// TIA Portal V20 export
Screen "Sew_APC"  1276x673
  ScreenItem "Rectangle_3" at 194,365 size 865x300  Type=HmiRectangle
  ScreenItem "Rectangle_1" at 195,113 size 866x250  Type=HmiRectangle
  ScreenItem "Title_ScreenOverview_X390_Y2" at 390,7 size 510x57  Type=HmiTextBox
  ScreenItem "符号 IO 域_7" at 479,72 size 290x38  Type=HmiSymbolicIOField
  ScreenItem "Text field_1" at 194,113 size 866x31  Type=HmiTextBox
  ScreenItem "按钮_2" at 279,171 size 140x60  Type=HmiButton
  ScreenItem "permanentareaborderrectangle" at 0,0 size 0x0  Type=HmiRectangle
  ScreenItem "Line_Header_X0_Y64" at 0,65 size 1276x0  Type=HmiLine
  ScreenItem "Button_Back" at 2,2 size 90x60  Type=HmiButton
  ScreenItem "Frame_SendToDrive_1" at 201,369 size 199x294  Type=HmiRectangle
  ScreenItem "Text_ConrolDataToDrive_1" at 205,373 size 148x21  Type=HmiTextBox
  ScreenItem "Text_DigitalOutputs_33" at 229,397 size 146x16  Type=HmiTextBox
  ScreenItem "Text_DigitalOutputs_34" at 229,412 size 124x16  Type=HmiTextBox
  ScreenItem "Text_DigitalOutputs_35" at 229,428 size 124x16  Type=HmiTextBox
  ScreenItem "Text_DigitalOutputs_40" at 229,444 size 124x16  Type=HmiTextBox
  ScreenItem "Text_DigitalOutputs_36" at 229,460 size 124x16  Type=HmiTextBox
  ScreenItem "Text_DigitalOutputs_37" at 229,476 size 124x16  Type=HmiTextBox
  ScreenItem "Text_DigitalOutputs_24" at 229,492 size 124x16  Type=HmiTextBox
  ScreenItem "Text_DigitalOutputs_38" at 229,508 size 124x16  Type=HmiTextBox
  ScreenItem "Text_DigitalOutputs_25" at 229,524 size 124x16  Type=HmiTextBox
  ScreenItem "Text_DigitalOutputs_39" at 229,540 size 124x16  Type=HmiTextBox
  ScreenItem "Text_DigitalOutputs_26" at 229,556 size 124x16  Type=HmiTextBox
  ScreenItem "Text_DigitalOutputs_1" at 229,572 size 124x16  Type=HmiTextBox
  ScreenItem "Text_DigitalOutputs_28" at 229,588 size 161x16  Type=HmiTextBox
  ScreenItem "Text_DigitalOutputs_30" at 229,604 size 124x16  Type=HmiTextBox
  ScreenItem "Text_DigitalOutputs_31" at 229,620 size 124x16  Type=HmiTextBox
  ScreenItem "Text_DigitalOutputs_32" at 229,636 size 124x16  Type=HmiTextBox
  ScreenItem "LED_1_Left_23" at 0,0 size 100x30  Type=HmiCircle
  ScreenItem "LED_1_Left_22" at 0,0 size 100x30  Type=HmiCircle
  ScreenItem "LED_1_Left_21" at 0,0 size 100x30  Type=HmiCircle
  ScreenItem "LED_1_Left_20" at 0,0 size 100x30  Type=HmiCircle
  ScreenItem "LED_1_Left_19" at 0,0 size 100x30  Type=HmiCircle
  ScreenItem "LED_1_Left_18" at 0,0 size 100x30  Type=HmiCircle
  ScreenItem "LED_1_Left_40" at 0,0 size 100x30  Type=HmiCircle
  ScreenItem "LED_1_Left_17" at 0,0 size 100x30  Type=HmiCircle
  ScreenItem "LED_1_Left_39" at 0,0 size 100x30  Type=HmiCircle
  ScreenItem "LED_1_Left_16" at 0,0 size 100x30  Type=HmiCircle
  ScreenItem "LED_1_Left_38" at 0,0 size 100x30  Type=HmiCircle
  ScreenItem "LED_1_Left_37" at 0,0 size 100x30  Type=HmiCircle
  ScreenItem "LED_1_Left_36" at 0,0 size 100x30  Type=HmiCircle
  ScreenItem "LED_1_Left_35" at 0,0 size 100x30  Type=HmiCircle
  ScreenItem "LED_1_Left_34" at 0,0 size 100x30  Type=HmiCircle
  ScreenItem "LED_1_Left_33" at 0,0 size 100x30  Type=HmiCircle
  ScreenItem "Frame_SendToDrive_3" at 405,369 size 199x294  Type=HmiRectangle
  ScreenItem "Text_ConrolDataToDrive_2" at 407,372 size 148x23  Type=HmiTextBox
  ScreenItem "Text_DigitalOutputs_2" at 426,395 size 124x20  Type=HmiTextBox
  ScreenItem "Text_DigitalOutputs_3" at 426,410 size 124x20  Type=HmiTextBox
  ScreenItem "Text_DigitalOutputs_4" at 426,426 size 124x20  Type=HmiTextBox
  ScreenItem "Text_DigitalOutputs_5" at 426,458 size 124x20  Type=HmiTextBox
  ScreenItem "Text_DigitalOutputs_6" at 426,474 size 124x20  Type=HmiTextBox
  ScreenItem "Text_DigitalOutputs_7" at 426,490 size 158x20  Type=HmiTextBox
  ScreenItem "Text_DigitalOutputs_8" at 426,506 size 124x20  Type=HmiTextBox
  ScreenItem "Text_DigitalOutputs_9" at 426,442 size 124x20  Type=HmiTextBox
  ScreenItem "Text_ConrolDataToDrive_3" at 407,372 size 148x23  Type=HmiTextBox
  ScreenItem "LED_1_Left_8" at 0,0 size 100x30  Type=HmiCircle
  ScreenItem "LED_1_Left_7" at 0,0 size 100x30  Type=HmiCircle
  ScreenItem "LED_1_Left_6" at 0,0 size 100x30  Type=HmiCircle
  ScreenItem "LED_1_Left_5" at 0,0 size 100x30  Type=HmiCircle
  ScreenItem "LED_1_Left_4" at 0,0 size 100x30  Type=HmiCircle
  ScreenItem "LED_1_Left_3" at 0,0 size 100x30  Type=HmiCircle
  ScreenItem "LED_1_Left_2" at 0,0 size 100x30  Type=HmiCircle
  ScreenItem "LED_1_Left_1" at 0,0 size 100x30  Type=HmiCircle
  ScreenItem "Text_DigitalOutputs_10" at 426,522 size 124x20  Type=HmiTextBox
  ScreenItem "Text_DigitalOutputs_11" at 426,538 size 124x20  Type=HmiTextBox
  ScreenItem "Text_DigitalOutputs_12" at 426,554 size 124x20  Type=HmiTextBox
  ScreenItem "Text_DigitalOutputs_13" at 426,586 size 158x20  Type=HmiTextBox
  ScreenItem "Text_DigitalOutputs_14" at 426,602 size 124x20  Type=HmiTextBox
  ScreenItem "Text_DigitalOutputs_15" at 426,618 size 158x20  Type=HmiTextBox
  ScreenItem "Text_DigitalOutputs_16" at 426,634 size 124x20  Type=HmiTextBox
  ScreenItem "Text_DigitalOutputs_17" at 426,570 size 186x20  Type=HmiTextBox
  ScreenItem "LED_1_Left_9" at 0,0 size 100x30  Type=HmiCircle
  ScreenItem "LED_1_Left_10" at 0,0 size 100x30  Type=HmiCircle
  ScreenItem "LED_1_Left_11" at 0,0 size 100x30  Type=HmiCircle
  ScreenItem "LED_1_Left_12" at 0,0 size 100x30  Type=HmiCircle
  ScreenItem "LED_1_Left_13" at 0,0 size 100x30  Type=HmiCircle
  ScreenItem "LED_1_Left_14" at 0,0 size 100x30  Type=HmiCircle
  ScreenItem "LED_1_Left_15" at 0,0 size 100x30  Type=HmiCircle
  ScreenItem "LED_1_Left_24" at 0,0 size 100x30  Type=HmiCircle
  ScreenItem "Text field_3" at 194,308 size 868x31  Type=HmiTextBox
  ScreenItem "Text field_8" at 622,447 size 94x29  Type=HmiTextBox
  ScreenItem "FaultNo" at 724,446 size 65x31  Type=HmiIOField
  ScreenItem "Text field_2" at 622,411 size 94x29  Type=HmiTextBox
  ScreenItem "FaultNo_2" at 724,410 size 65x31  Type=HmiIOField
  ScreenItem "Text field_4" at 622,375 size 94x29  Type=HmiTextBox
  ScreenItem "FaultNo_3" at 724,374 size 65x31  Type=HmiIOField
  ScreenItem "Graphic view_1" at 698,-47 size 128x565  Type=HmiGraphicView
